(* IEC 61131-3 sources: botanik2/src/libbotanik/plc/blocks, 6 files *)

(* ---- actuator.st ---- *)
(* Open/close coil pairs, driven to a fractional target by timing
   ------------------------------------------------------------------------ *)

(* Drives an open/close coil pair to a fractional target by TIMING the strokes.
   No position feedback: the position is an ESTIMATE, a stroke to either end
   runs SEAT_MS extra to re-datum, and it is UNKNOWN until one has.

   Three invariants: the coils are never both energised, a reversal always
   passes through REVERSE_MS with both dropped (a contactor that makes before
   the other breaks shorts the motor), and a move under MIN_RUN_MS is not made
   at all. *)

FUNCTION ACT_WANT : USINT
(* The direction TGT asks for: 0 none, 1 open, 2 close. *)
VAR_INPUT
  MODE : USINT;
  P    : REAL;
  TGT  : REAL;
  DB   : REAL;
END_VAR
VAR
  err : REAL;
END_VAR
  IF MODE = 0 THEN
    (* Nothing is known about where it sits, so there is no error to compute:
       drive to whichever end the target is nearer, and datum there. *)
    IF TGT >= 1.0 - DB THEN ACT_WANT := 1; ELSE ACT_WANT := 2; END_IF;
  ELSE
    err := TGT - P;
    IF   err >  DB       THEN ACT_WANT := 1;
    ELSIF err < -DB THEN ACT_WANT := 2;
    ELSE ACT_WANT := 0;
    END_IF;
  END_IF;
END_FUNCTION

FUNCTION_BLOCK ACTUATOR
VAR_INPUT
  TARGET       : REAL;    (* 0 closed .. 1 open; clamped *)
  OPEN_MS      : UDINT;
  CLOSE_MS     : UDINT;
  SEAT_MS      : UDINT;   (* extra run at an end, to re-datum. Safe because
                             the drive has a limit switch: it cuts the
                             motor, so the over-run costs nothing *)
  MIN_RUN_MS   : UDINT;
  REVERSE_MS   : UDINT;
  DB           : REAL;    (* how far off target is close enough *)
  REDATUM      : REAL;    (* full strokes between datums; 0 disables *)
  HOLD         : BOOL;    (* this one does not have the bus this scan: keep
                             the clock, decide nothing. A target of "stay"
                             would still send an unknown one to datum. *)
  PRESET_KNOWN : BOOL;    (* the first scan finds it at PRESET_POS *)
  PRESET_POS   : REAL;
  NOW          : UDINT;   (* sys_now_ms: the scan clock, not an elapsed time *)
END_VAR
VAR_OUTPUT
  OPEN_CMD  : BOOL;
  CLOSE_CMD : BOOL;    (* never true at the same time as OPEN_CMD *)
  POS       : REAL;    (* only meaningful once KNOWN *)
  KNOWN     : BOOL;
  MOVING    : BOOL;
  STATE     : USINT;   (* 0 UNKNOWN 1 CLOSING 2 CLOSED 3 OPENING 4 OPEN *)
  DRIFT     : REAL;    (* travel since the last datum, in full strokes. No
                          drive reports a fault, so this is the only wear
                          signal there is - it is published for a person *)
END_VAR
VAR
  p       : REAL;
  run_ms  : UDINT;
  wait_ms : UDINT;
  mode    : USINT;
  dir     : USINT;   (* 0 none, 1 open, 2 close *)
  seating : BOOL;    (* this stroke ends at a seat, so snap there *)
  datum   : BOOL;    (* ...and it is the one establishing position *)
  moved   : REAL;
  pending : REAL := -1.0;   (* where to go once the detour finishes, or -1 *)
  last    : UDINT;
  seeded  : BOOL := FALSE;
END_VAR
VAR_TEMP
  elapsed   : UDINT;
  tgt       : REAL;
  ran       : UDINT;
  span      : UDINT;
  delta     : REAL;
  want      : USINT;
  partial   : BOOL;
  is_datum  : BOOL;
  to_end    : BOOL;
  distance  : REAL;
  stroke_ms : UDINT;
  commit    : BOOL;
END_VAR
  IF seeded THEN
    elapsed := NOW - last;
  ELSE
    elapsed := 0;
    seeded  := TRUE;
    (* Position known without a datum stroke, only where the wiring
       establishes it: the screen deploys on the de-energised coil, so a
       controller that was not driving anything left the fabric out. *)
    IF PRESET_KNOWN THEN
      p := LIMIT(0.0, PRESET_POS, 1.0);
      IF p <= 0.0 THEN mode := 2; ELSE mode := 4; END_IF;
    END_IF;
  END_IF;
  last := NOW;

  IF NOT HOLD THEN

    tgt := LIMIT(0.0, TARGET, 1.0);

    (* A re-datum detour owns the target for the WHOLE scan: the mid-stroke
       interrupt below sees the caller's target pointing the other way, and
       would abort the detour on the next scan. *)
    IF pending >= 0.0 THEN
      IF mode = 2 THEN
        tgt     := pending;
        pending := -1.0;
      ELSE
        tgt := 0.0;
      END_IF;
    END_IF;

    IF run_ms > 0 THEN
      (* Only the part of this scan the coil was actually energised for counts as
         travel; the rest belongs to the next decision. *)
      IF elapsed < run_ms THEN ran := elapsed; ELSE ran := run_ms; END_IF;
      IF dir = 1 THEN span := OPEN_MS; ELSE span := CLOSE_MS; END_IF;
      (* A zero travel time is a misconfiguration: treat it as instant. *)
      IF span > 0 THEN delta := UDINT_TO_REAL(ran) / UDINT_TO_REAL(span);
      ELSE delta := 1.0;
      END_IF;
      (* Every stroke adds to the uncertainty, whichever way it went; only
         reaching a stop takes it back. *)
      moved := moved + delta;
      IF dir = 1 THEN p := LIMIT(0.0, p + delta, 1.0);
      ELSE            p := LIMIT(0.0, p - delta, 1.0);
      END_IF;
      run_ms := run_ms - ran;

      IF run_ms = 0 THEN
        (* The stroke ran past the mechanical stop, so the estimate is a fact
           rather than an integration. *)
        IF seating THEN
          IF dir = 1 THEN p := 1.0; ELSE p := 0.0; END_IF;
          moved := 0.0;
        END_IF;
        dir     := 0;
        seating := FALSE;
        datum   := FALSE;
        (* Dead time after EVERY stroke, not only an interrupted one: the move
           that follows one which just seated can only be the opposite
           direction, and it would otherwise start in this very scan. *)
        wait_ms := REVERSE_MS;
        IF p <= 0.0 THEN mode := 2; ELSE mode := 4; END_IF;
      ELSIF NOT datum THEN
        (* The target moved the other way mid-stroke. A stroke is otherwise
           COMMITTED - a seating run must be allowed to overrun the estimate,
           which is the whole point of it - so only the opposite direction
           interrupts, never "we are close enough now". *)
        want := ACT_WANT(MODE := mode, P := p, TGT := tgt, DB := DB);
        IF want <> 0 AND want <> dir THEN
          run_ms  := 0;
          seating := FALSE;
          dir     := 0;
          wait_ms := REVERSE_MS;
          IF p <= 0.0 THEN mode := 2; ELSE mode := 4; END_IF;
        END_IF;
      END_IF;
    ELSIF wait_ms > 0 THEN
      IF wait_ms > elapsed THEN wait_ms := wait_ms - elapsed; ELSE wait_ms := 0; END_IF;
    END_IF;

    IF run_ms = 0 AND wait_ms = 0 THEN
      want := ACT_WANT(MODE := mode, P := p, TGT := tgt, DB := DB);
      (* Nothing is wanted, so nothing happens - INCLUDING a re-datum. Letting
         one fire on a steady target would send the actuator to the seat and back
         while nobody asked it to move at all. *)
      IF want <> 0 THEN
        (* Only for a move that ENDS PARTWAY. One to either end runs onto the
           stop and re-datums by itself, so a detour would be a wasted stroke. *)
        partial := tgt > DB AND tgt < 1.0 - DB;
        IF pending < 0.0 AND REDATUM > 0.0 AND moved >= REDATUM
           AND mode <> 0 AND partial THEN
          pending := tgt;
          tgt     := 0.0;
          (* Recomputed: deciding the direction from the caller's target and then
             redirecting the stroke would drive the wrong way. *)
          want := ACT_WANT(MODE := mode, P := p, TGT := tgt, DB := DB);
          IF want = 0 THEN pending := -1.0; END_IF;
        END_IF;

        IF want <> 0 THEN
          is_datum := mode = 0;
          to_end   := is_datum OR tgt <= DB OR tgt >= 1.0 - DB;
          IF want = 1 THEN span := OPEN_MS; ELSE span := CLOSE_MS; END_IF;
          (* A datum stroke assumes the worst case, a full travel away. *)
          IF is_datum THEN distance := 1.0; ELSE distance := tgt - p; END_IF;
          distance := ABS(distance);
          stroke_ms := REAL_TO_UDINT(distance * UDINT_TO_REAL(span));
          commit  := TRUE;
          IF to_end THEN
            stroke_ms := stroke_ms + SEAT_MS;      (* overrun onto the stop, re-datuming *)
          ELSIF stroke_ms < MIN_RUN_MS THEN
            commit := FALSE;               (* not worth a twitch *)
          END_IF;
          IF commit THEN
            IF stroke_ms = 0 THEN stroke_ms := 1; END_IF;   (* always make progress *)
            dir     := want;
            run_ms  := stroke_ms;
            seating := to_end;
            datum   := is_datum;
            IF want = 1 THEN mode := 3; ELSE mode := 1; END_IF;
          END_IF;
        END_IF;
      END_IF;
    END_IF;
  END_IF;

  OPEN_CMD  := dir = 1 AND run_ms > 0;
  CLOSE_CMD := dir = 2 AND run_ms > 0;
  MOVING    := OPEN_CMD OR CLOSE_CMD;
  POS       := p;
  KNOWN     := mode <> 0;
  STATE     := mode;
  DRIFT     := moved;
END_FUNCTION_BLOCK

(* ---- analog.st ---- *)
(* Analog conditioning: a latch, a three-step ladder, a deadband, a DC rail
   ------------------------------------------------------------------------ *)

(* Latches ON at its rising edge and OFF below the falling one, holding
   between the two: a reading sitting on a threshold decides once. *)
FUNCTION_BLOCK BAND_LATCH
VAR_INPUT
  IN   : REAL;
  RISE : REAL;   (* engages at or above *)
  FALL : REAL;   (* releases at or below *)
END_VAR
VAR_OUTPUT
  Q : BOOL;
END_VAR
  IF   IN >= RISE THEN Q := TRUE;
  ELSIF IN <= FALL THEN Q := FALSE;
  END_IF;
END_FUNCTION_BLOCK

(* Three rungs, each holding its OWN release band. All three are evaluated: a
   rung that stopped being asked keeps whichever side of itself the reading
   was last on. *)
FUNCTION_BLOCK STAIRCASE3
VAR_INPUT
  IN   : REAL;
  LO   : REAL;
  MED  : REAL;
  HI   : REAL;
  HYST : REAL;
END_VAR
VAR_OUTPUT
  Q : USINT;
END_VAR
VAR
  rung1 : BAND_LATCH;
  rung2 : BAND_LATCH;
  rung3 : BAND_LATCH;
END_VAR
VAR_TEMP
  h : REAL;
END_VAR
  (* A negative hysteresis is no hysteresis, never an inverted band. *)
  IF HYST < 0.0 THEN h := 0.0; ELSE h := HYST; END_IF;

  rung1(IN := IN, RISE := LO,  FALL := LO  - h);
  rung2(IN := IN, RISE := MED, FALL := MED - h);
  rung3(IN := IN, RISE := HI,  FALL := HI  - h);

  Q := 0;
  IF rung1.Q THEN Q := 1; END_IF;
  IF rung2.Q THEN Q := 2; END_IF;
  IF rung3.Q THEN Q := 3; END_IF;
END_FUNCTION_BLOCK

FUNCTION_BLOCK DEADBAND
(* Report a value only once it has MOVED more than BAND, so a reading that
   twitches in its last digit does not cost a status write per scan. Cold, the
   first reading is reported whatever it is rather than suppressed against a
   held value from before the gap. *)
VAR_INPUT
  V    : REAL;
  BAND : REAL;
END_VAR
VAR_OUTPUT
  Y : REAL;
END_VAR
VAR
  held : REAL;
  seeded : BOOL := FALSE;
END_VAR
VAR_TEMP
  diff : REAL;
END_VAR
  diff := V - held;
  IF NOT seeded OR ABS(diff) > BAND THEN
    held   := V;
    seeded := TRUE;
  END_IF;
  Y := held;
END_FUNCTION_BLOCK

FUNCTION_BLOCK DC_RAIL
(* One DC rail off a divider: averaged, then deadbanded. The first says what
   the rail is doing, the second says when that is worth a status write. *)
VAR_INPUT
  V      : REAL;
  V_Q    : QUALITY;
  LO     : REAL;    (* the floor the rail is judged against *)
  AVG_MS : UINT;
  BAND   : REAL;
  NOW    : UDINT;   (* sys_now_ms: the scan clock, not an elapsed time *)
END_VAR
VAR_OUTPUT
  Y       : REAL;
  Q       : QUALITY;
  HEALTHY : BOOL;
END_VAR
VAR
  avg : EWMA;
  db  : DEADBAND;
  seen : BOOL := FALSE;
END_VAR
  (* Only a MEASURED sample is folded in: the row reads its declared value
     while the bus is coming up, and folding that seeds the average at zero,
     so the rail reads under its floor until the filter climbs out - a supply
     alarm on every boot. CALLED either way, since the filter reads the clock.
     The band is left open: LO is what HEALTHY is judged against, not a clamp. *)
  avg.X     := V;
  avg.Q_IN  := V_Q;
  avg.TAU_S := UINT_TO_REAL(AVG_MS) / 1000.0;
  avg.NOW   := NOW;
  avg.LO    := 0.0;
  avg.HI    := 0.0;
  avg();
  IF GOOD(V_Q) THEN
    db(V := avg.Y, BAND := BAND);
    seen := TRUE;
  END_IF;
  (* A rail nobody is measuring has no voltage to publish. Its LAST average
     stays in the filter, so a divider that comes back rejoins where it left. *)
  Y := db.Y;
  Q := avg.Q;

  (* A divider that has NEVER answered is the bus still coming up. One that has
     answered and then stopped is a rail nobody can see, which is a fault. *)
  IF GOOD(V_Q) THEN HEALTHY := avg.Y >= LO;
  ELSE              HEALTHY := NOT seen;
  END_IF;
END_FUNCTION_BLOCK

(* ---- filters.st ---- *)
(* The one filter every measured row is published through
   ------------------------------------------------------------------------ *)

FUNCTION_BLOCK EWMA
(* An exponentially-weighted moving average of X, clamped to the row's band,
   and the verdict on whether this beat had anything to average. *)
VAR_INPUT
  X     : REAL;
  Q_IN  : QUALITY;   (* what fed X this beat is worth *)
  TAU_S : REAL;
  NOW   : UDINT;     (* sys_now_ms: the scan clock, not an elapsed time *)
  LO    : REAL;      (* the published band; HI <= LO publishes unclamped *)
  HI    : REAL;
END_VAR
VAR_OUTPUT
  Y : REAL;
  (* Q_GOOD this beat measured it; Q_HELD it holds an average of readings it
     did measure; Q_NONE nothing has ever fed it, so Y is the band's floor. *)
  Q : QUALITY;
END_VAR
VAR
  avg  : REAL;
  last : UDINT;
  primed : BOOL := FALSE;
END_VAR
VAR_TEMP
  dt_s  : REAL;
  alpha : REAL;
END_VAR
  (* Call it every scan and say so with Q_IN, rather than skipping it while
     the reading is out: skipped, the first sample after the outage arrives
     with the whole outage as its interval and the average SNAPS to it instead
     of rejoining where it left. Five minutes against a 30 s tau is alpha 0.91. *)
  Q := QUAL(GOOD(Q_IN), primed);
  IF NOT GOOD(Q_IN) THEN
    last := NOW;
    (* Primed, Y keeps the last average and Q says nothing measured it this
       beat. Never primed, nothing has EVER measured this: the band's floor
       rather than a default zero, which on a temperature reads like a
       measurement of a freezing house. *)
    IF NOT primed THEN Y := LO; END_IF;
    RETURN;
  END_IF;

  IF NOT primed THEN
    (* Starts AT its first reading rather than climbing to it from zero. The
       clock is adopted with it, so the first real interval is the second
       scan's and never the time since boot. *)
    avg    := X;
    primed := TRUE;
  ELSIF TAU_S <= 0.0 THEN
    avg := X;
  ELSE
    dt_s  := UDINT_TO_REAL(NOW - last) / 1000.0;
    alpha := dt_s / (TAU_S + dt_s);
    avg   := avg + alpha * (X - avg);
  END_IF;
  last := NOW;

  IF HI > LO THEN Y := LIMIT(LO, avg, HI); ELSE Y := avg; END_IF;
END_FUNCTION_BLOCK

(* ---- meter.st ---- *)
(* Integrating a rate, and differentiating a quantity
   ------------------------------------------------------------------------ *)

(* HOLD is "keep the clock, count nothing": see EWMA for why a clocked block
   needs one rather than being skipped. *)

FUNCTION_BLOCK INTEGRAL
(* Count RATE for as long as it has been in force. Needs the REAL elapsed: a
   program that ran 400 ms late delivered 400 ms of water. *)
VAR_INPUT
  RATE_PER_S : REAL;
  CUTOFF     : REAL;   (* below this the rate counts as zero *)
  HOLD       : BOOL;
  SEED       : REAL;   (* the total the FIRST scan starts from: a retained row
                          carries what was metered before this run, and a
                          totaliser that restarts at zero unmakes it *)
  NOW        : UDINT;
END_VAR
VAR_OUTPUT
  TOTAL : REAL;
  RATE  : REAL;   (* the rate actually counted, after the cutoff *)
END_VAR
VAR
  last : UDINT;
  seeded : BOOL := FALSE;
END_VAR
VAR_TEMP
  elapsed : UDINT;
  r       : REAL;
END_VAR
  IF seeded THEN
    elapsed := NOW - last;
  ELSE
    elapsed := 0;
    seeded  := TRUE;
    TOTAL   := SEED;
  END_IF;
  last := NOW;

  IF NOT HOLD THEN
    r := RATE_PER_S;
    (* A meter idling on noise must not total a plausible volume with the pump
       off, so anything inside the cutoff counts as nothing at all. *)
    IF CUTOFF > 0.0 AND ABS(r) < CUTOFF THEN r := 0.0; END_IF;
    RATE  := r;
    TOTAL := TOTAL + r * (UDINT_TO_REAL(elapsed) / 1000.0);
  END_IF;
END_FUNCTION_BLOCK

FUNCTION_BLOCK DERIVATIVE
(* The rate a quantity is changing at, over a WINDOW rather than per scan: a
   pulse meter counts in whole litres, so scan to scan it reads either zero or
   one pulse's worth and never the flow. *)
VAR_INPUT
  QUANTITY  : REAL;
  WINDOW_MS : UDINT;   (* 0 differentiates every scan *)
  PRESET    : BOOL;    (* adopt QUANTITY without reporting a rate *)
  NOW       : UDINT;
END_VAR
VAR_OUTPUT
  RATE : REAL;   (* per second; the last COMPLETED window, held between them *)
END_VAR
VAR
  prev   : REAL;
  window : UDINT;   (* time accumulated into this window *)
  last   : UDINT;
  seeded  : BOOL := FALSE;
END_VAR
VAR_TEMP
  elapsed : UDINT;
END_VAR
  IF seeded THEN elapsed := NOW - last;
  ELSE elapsed := 0;
  END_IF;
  last := NOW;

  IF PRESET OR NOT seeded THEN
    (* Adopt the reading rather than differencing against a zero: the first
       window would otherwise report the whole counter as a rate. *)
    prev   := QUANTITY;
    window := 0;
    seeded := TRUE;
    RATE   := 0.0;
  ELSE
    window := window + elapsed;
    IF window > 0 AND window >= WINDOW_MS THEN
      (* Over the time actually accumulated, not the nominal window: a late
         scan overshoots it, and the nominal figure would report a rate that
         never happened. *)
      RATE   := (QUANTITY - prev) / (UDINT_TO_REAL(window) / 1000.0);
      prev   := QUANTITY;
      window := 0;
    END_IF;
  END_IF;
END_FUNCTION_BLOCK

(* ---- pid.st ---- *)
(* The PID loop
   ------------------------------------------------------------------------ *)

FUNCTION_BLOCK PID
(* Holds a reading at a setpoint. Direct-acting by default: the output rises as
   the reading FALLS (heating, filling). Three departures from the textbook sum,
   all affecting tuning: derivative on the MEASUREMENT, so a typed setpoint does
   not slam the output; conditional integration, so there is no back-calculation
   gain to tune; and the integral clamped to the output SPAN, not its limits.

   RESET clears the history in place - the loop still runs this scan, on a cold
   integral. That is what a law does when it stops being able to see the plant:
   effort wound up against a house nobody is measuring is a claim about a past
   the loop no longer has. *)
VAR_INPUT
  SP      : REAL;
  PV      : REAL;
  KP      : REAL;
  KI      : REAL;    (* per (error x second); 0 is NO integral action *)
  KD      : REAL;
  OUT_MIN : REAL;
  OUT_MAX : REAL;
  D_TAU_S : REAL;    (* derivative lowpass; 0 is unfiltered *)
  REVERSE : BOOL;    (* output rises as the reading does *)
  RESET   : BOOL;
  NOW     : UDINT;   (* sys_now_ms: the scan clock, not an elapsed time *)
END_VAR
VAR_OUTPUT
  Y         : REAL;
  ERR       : REAL;   (* sign-corrected: positive asks for more output *)
  INTEGRAL  : REAL;   (* in OUTPUT units - what to watch when a loop misbehaves *)
  SATURATED : BOOL;
END_VAR
VAR
  last    : UDINT;
  seeded  : BOOL := FALSE;
  prev_pv : REAL;
  deriv   : REAL;
END_VAR
VAR_TEMP
  dt_s      : REAL;
  d_raw     : REAL;
  alpha     : REAL;
  p_term    : REAL;
  d_term    : REAL;
  trial     : REAL;
  winding   : BOOL;
  unclamped : REAL;
  i_lo      : REAL;
  i_hi      : REAL;
END_VAR
  IF RESET THEN
    INTEGRAL := 0.0;
    prev_pv  := 0.0;
    deriv    := 0.0;
    seeded   := FALSE;
  END_IF;

  (* The first scan adopts the reading, so the derivative starts at zero rather
     than at PV/dt, which is a very large number. *)
  IF seeded THEN
    dt_s := UDINT_TO_REAL(NOW - last) / 1000.0;
  ELSE
    dt_s      := 0.0;
    prev_pv := PV;
    seeded  := TRUE;
  END_IF;
  last := NOW;

  IF REVERSE THEN ERR := PV - SP; ELSE ERR := SP - PV; END_IF;

  IF dt_s > 0.0 THEN
    d_raw := (PV - prev_pv) / dt_s;
    IF D_TAU_S > 0.0 THEN
      alpha := dt_s / (D_TAU_S + dt_s);
      deriv := deriv + alpha * (d_raw - deriv);
    ELSE
      deriv := d_raw;
    END_IF;
    prev_pv := PV;
  END_IF;

  (* Derivative on the measurement opposes the reading's movement, so it enters
     with the sign the action gives it. *)
  p_term := KP * ERR;
  IF REVERSE THEN d_term := KD * deriv; ELSE d_term := -(KD * deriv); END_IF;

  IF KI = 0.0 THEN
    (* No integral ACTION means no integral TERM, not a frozen one: KI is
       operator-editable, and whatever had accumulated would go on commanding
       the output for ever with nothing able to remove it. *)
    INTEGRAL := 0.0;
  ELSIF dt_s > 0.0 THEN
    (* Conditional integration: only when it does not push further into a limit
       the output is already against. *)
    trial := p_term + INTEGRAL + d_term;
    winding := (trial >= OUT_MAX AND ERR > 0.0)
            OR (trial <= OUT_MIN AND ERR < 0.0);
    IF NOT winding THEN
      INTEGRAL := INTEGRAL + KI * ERR * dt_s;
      (* Clamped so the integral can SPAN the output, NOT to the output's own
         limits: with a non-zero floor, LIMIT(20, i, 100) would clamp a fresh
         integral of 0.01 UP to 20 and the winding test would pin it there for
         good. Zero has to stay reachable from either side. *)
      IF OUT_MIN < 0.0 THEN i_lo := OUT_MIN; ELSE i_lo := 0.0; END_IF;
      IF OUT_MAX > 0.0 THEN i_hi := OUT_MAX; ELSE i_hi := 0.0; END_IF;
      INTEGRAL := LIMIT(i_lo, INTEGRAL, i_hi);
    END_IF;
  END_IF;

  unclamped   := p_term + INTEGRAL + d_term;
  SATURATED := (unclamped > OUT_MAX) OR (unclamped < OUT_MIN);
  Y         := LIMIT(OUT_MIN, unclamped, OUT_MAX);
END_FUNCTION_BLOCK

(* ---- timers.st ---- *)
(* The two dwell timers: off-delay and on-delay, in milliseconds
   ------------------------------------------------------------------------ *)

(* Off-delay: true while IN is, and for PT after it drops. An overrun - "keep
   the roof shut for a quarter of an hour after the last drop". *)
FUNCTION_BLOCK TOF_MS
VAR_INPUT
  IN  : BOOL;
  PT  : UDINT;   (* ms *)
  NOW : UDINT;   (* sys_now_ms: the scan clock, not an elapsed time *)
END_VAR
VAR_OUTPUT
  Q  : BOOL;
  ET : UDINT;
END_VAR
VAR
  (* Measured from when this timer last ran, so a scan it missed costs it
     nothing. *)
  last : UDINT;
  seeded : BOOL := FALSE;
END_VAR
VAR_TEMP
  elapsed : UDINT;
END_VAR
  IF seeded THEN elapsed := NOW - last;
  ELSE elapsed := 0; seeded := TRUE;
  END_IF;
  last := NOW;

  IF IN THEN
    ET := 0;
    Q  := TRUE;
  ELSIF Q THEN
    (* Saturating, so a scan that arrives after PT cannot wrap the counter. *)
    IF ET > UDINT#4000000000 - elapsed THEN ET := UDINT#4000000000;
    ELSE ET := ET + elapsed;
    END_IF;
    IF ET >= PT THEN Q := FALSE; END_IF;
  END_IF;
END_FUNCTION_BLOCK

FUNCTION_BLOCK TON_MS
(* On-delay: true once IN has held true for PT, false the moment it drops.
   A dwell - "has been wet for 30 s", "has been silent long enough to alarm". *)
VAR_INPUT
  IN  : BOOL;
  PT  : UDINT;   (* ms *)
  NOW : UDINT;   (* sys_now_ms: the scan clock, not an elapsed time *)
END_VAR
VAR_OUTPUT
  Q  : BOOL;
  ET : UDINT;
END_VAR
VAR
  last : UDINT;
  seeded : BOOL := FALSE;
END_VAR
VAR_TEMP
  elapsed : UDINT;
END_VAR
  IF seeded THEN elapsed := NOW - last;
  ELSE elapsed := 0; seeded := TRUE;
  END_IF;
  last := NOW;

  IF NOT IN THEN
    ET := 0;
    Q  := FALSE;
  ELSE
    (* Saturating, so a scan that arrives after PT cannot wrap the counter. *)
    IF ET > UDINT#4000000000 - elapsed THEN ET := UDINT#4000000000;
    ELSE ET := ET + elapsed;
    END_IF;
    Q := ET >= PT;
  END_IF;
END_FUNCTION_BLOCK
